FUNCTION_BLOCK Valvula_Solenoide_HMI (* Service Interface Function Block Type *)
  (* Standard: 61499-2 *)
  (* Version 1.0, 04/11/2026, Hidryco, Hidryco, IHM da Valvula_Solenoide (tags da IO List da Nereda) *)
  PACKAGE Hidryco.HidrycoLib;
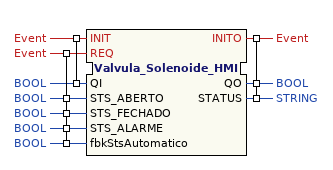
  EVENT_INPUT
    INIT WITH QI;
    REQ WITH STS_ABERTO, STS_FECHADO, STS_ALARME, fbkStsAutomatico; (* Atualizacao de status *)
  END_EVENT
  EVENT_OUTPUT
    INITO WITH QO, STATUS;
  END_EVENT
  VAR_INPUT
    QI : BOOL;
    STS_ABERTO : BOOL; (* Valvula aberta *)
    STS_FECHADO : BOOL; (* Valvula fechada *)
    STS_ALARME : BOOL; (* Discrepancia entre comando e fim de curso *)
    fbkStsAutomatico : BOOL; (* Modo automatico (sempre FALSE: SV so manual) *)
  END_VAR
  VAR_OUTPUT
    QO : BOOL; (* Event Output Qualifier *)
    STATUS : STRING; (* Service Status *)
  END_VAR
  SERVICE /
    SEQUENCE 
    END_SEQUENCE
  END_SERVICE
END_FUNCTION_BLOCK
